// TIA Portal V19 export
// export: Created 2026-10-15T10:10:34.0661054Z, ExportSetting WithDefaults, DisplayName Totally Integrated Automation Portal, DisplayVersion V19, DisplayName TIA Portal Openness, DisplayVersion V19, DisplayName TIA Portal Version Control Interface, DisplayVersion V19, DisplayName STEP 7 Professional, DisplayVersion V19, DisplayName STEP 7 Safety, DisplayVersion V19, DisplayName WinCC Basic/Comfort/Advanced, DisplayVersion V19, DisplayName WinCC Unified, DisplayVersion V19
DATA_BLOCK "ROLL_Recipe1"   // DB6
{ S7_Optimized_Access := 'TRUE' }
VERSION : 0.1
// stored: AutoNumber true, DBAccessibleFromOPCUA true, DBAccessibleFromWebserver true, IsOnlyStoredInLoadMemory false, IsRetainMemResEnabled false, IsWriteProtectedInAS false, MemoryReserve 100
   VAR RETAIN
      DW : Array[0..41] of Word;
   END_VAR
BEGIN
   DW[5] := WORD#16#2360;
   DW[9] := WORD#16#2090;
   DW[13] := WORD#16#0001;
   DW[17] := WORD#16#2240;
   DW[21] := WORD#16#2060;
   DW[25] := WORD#16#2300;
   DW[29] := WORD#16#2120;
   DW[33] := WORD#16#2400;
   DW[37] := WORD#16#0001;
END_DATA_BLOCK
